(* IEC 61131-3 sources: plc-st-coding-agent/progress/evidence/f14_v14_remaining_20261113/jobs/codex_deepseek-v4pro (part 5) *)

(* ---- self-medium-04.raw_candidate_01.st ---- *)
FUNCTION_BLOCK FB
VAR_INPUT
    startBtn   : BOOL;
    resetBtn   : BOOL;
    doneSensor : BOOL;
    targetVol  : REAL;
    flowVol    : REAL;
END_VAR
VAR_OUTPUT
    valveOpen  : BOOL;
    fillsToday : INT;
END_VAR
VAR
    prevStartBtn   : BOOL := FALSE;
    prevResetBtn   : BOOL := FALSE;
    prevValveOpen  : BOOL := FALSE;
    pendingConfirm : BOOL := FALSE;
    accumulatedVol : REAL := 0.0;
    tmp_risingReset : BOOL;
    tmp_risingStart : BOOL;
    tmp_isFilling   : BOOL;
END_VAR

(* ENGINEERING_CONTRACT
   valveOpen: set only on start edge from idle/wait (R2,S2); holds while
             accumulatedVol < targetVol (R3,S9); closes on reset or target reach (R1,R3,S5).
   pendingConfirm: set same scan as target close; persists until confirmation,
             next start, or reset; sensor TRUE does not repeat count (R3-R5,S11).
   fillsToday: increments once on doneSensor with pending; saturates at 32767
             and still clears pending; reset zeros in same scan (R4-R5,S1,S6,S14).
   accumulatedVol: reset on reset/new bottle; adds flowVol only while filling,
             including start scan (R1-R3,S12).
   Priority: reset > start/new-bottle cancellation > flow/threshold close > done confirm.
   Units: targetVol/flowVol in mL REAL; fillsToday signed INT bounds 0..32767.
*)

(* CONTRACT_RULES [] *)

tmp_risingReset := resetBtn AND NOT prevResetBtn;
tmp_risingStart := startBtn AND NOT prevStartBtn;

IF tmp_risingReset THEN
    valveOpen      := FALSE;
    fillsToday     := 0;
    accumulatedVol := 0.0;
    pendingConfirm := FALSE;
ELSE
    tmp_isFilling := FALSE;

    IF tmp_risingStart AND NOT valveOpen THEN
        pendingConfirm := FALSE;
        accumulatedVol := 0.0;
        valveOpen      := TRUE;
        tmp_isFilling   := TRUE;
    ELSIF valveOpen THEN
        tmp_isFilling := TRUE;
    END_IF;

    IF tmp_isFilling THEN
        accumulatedVol := accumulatedVol + flowVol;
        IF accumulatedVol >= targetVol THEN
            valveOpen      := FALSE;
            pendingConfirm := TRUE;
            tmp_isFilling   := FALSE;
        END_IF;
    END_IF;

    IF pendingConfirm AND doneSensor THEN
        IF fillsToday < 32767 THEN
            fillsToday := fillsToday + 1;
        END_IF;
        pendingConfirm := FALSE;
    END_IF;
END_IF;

prevStartBtn  := startBtn;
prevResetBtn  := resetBtn;
prevValveOpen := valveOpen;

END_FUNCTION_BLOCK

(* ---- self-medium-05.candidate_01.st ---- *)
FUNCTION_BLOCK FB
VAR_INPUT
    enable : BOOL;
    resetBtn : BOOL;
    scanSeconds : LREAL;
    steamFlow : LREAL;
    fuelFlow : LREAL;
    steamTemp : LREAL;
    steamPressure : LREAL;
END_VAR
VAR_OUTPUT
    qualified : BOOL;
    dataFault : BOOL;
    qualifiedTon : LREAL;
    fuelTon : LREAL;
    revenue : LREAL;
    cost : LREAL;
    netProfit : LREAL;
END_VAR
VAR
    local_prev_reset : BOOL := FALSE;
    local_reset_edge : BOOL;
END_VAR

(* ENGINEERING_CONTRACT
   - qualified/dataFault: combinational, updated every scan.
   - qualifiedTon: accumulates only when enable, no fault, qualified, and no reset edge.
   - fuelTon: accumulates only when enable, no fault, and no reset edge.
   - resetBtn rising edge: clears both accumulators, higher priority than enable/fault.
   - reset is edge-only; held resetBtn does not repeatedly clear.
   - revenue/cost/netProfit recomputed every scan from current accumulators.
   - scanSeconds unit s, flows kg/s; both are legal under stated fault bounds.
*)

(* CONTRACT_RULES [] *)

local_reset_edge := resetBtn AND NOT local_prev_reset;

qualified := (steamTemp >= 447.0) AND (steamTemp <= 453.0)
             AND (steamPressure >= 3750.0) AND (steamPressure <= 3850.0);

dataFault := (scanSeconds <= 0.0)
             OR (scanSeconds > 10.0)
             OR (steamFlow < 0.0) OR (steamFlow > 90.0)
             OR (fuelFlow < 0.0) OR (fuelFlow > 6.0);

IF local_reset_edge THEN
    qualifiedTon := 0.0;
    fuelTon := 0.0;
ELSE
    IF enable AND NOT dataFault THEN
        fuelTon := fuelTon + (fuelFlow * scanSeconds / 1000.0);

        IF qualified THEN
            qualifiedTon := qualifiedTon + (steamFlow * scanSeconds / 1000.0);
        END_IF;
    END_IF;
END_IF;

revenue := qualifiedTon * 280.0;
cost := fuelTon * 1500.0;
netProfit := revenue - cost;

local_prev_reset := resetBtn;

END_FUNCTION_BLOCK

(* ---- self-medium-05.raw_candidate_01.st ---- *)
FUNCTION_BLOCK FB
VAR_INPUT
    enable : BOOL;
    resetBtn : BOOL;
    scanSeconds : LREAL;
    steamFlow : LREAL;
    fuelFlow : LREAL;
    steamTemp : LREAL;
    steamPressure : LREAL;
END_VAR
VAR_OUTPUT
    qualified : BOOL;
    dataFault : BOOL;
    qualifiedTon : LREAL;
    fuelTon : LREAL;
    revenue : LREAL;
    cost : LREAL;
    netProfit : LREAL;
END_VAR
VAR
    local_prev_reset : BOOL := FALSE;
    local_reset_edge : BOOL;
END_VAR

(* ENGINEERING_CONTRACT
   - qualified/dataFault: combinational, updated every scan.
   - qualifiedTon: accumulates only when enable, no fault, qualified, and no reset edge.
   - fuelTon: accumulates only when enable, no fault, and no reset edge.
   - resetBtn rising edge: clears both accumulators, higher priority than enable/fault.
   - reset is edge-only; held resetBtn does not repeatedly clear.
   - revenue/cost/netProfit recomputed every scan from current accumulators.
   - scanSeconds unit s, flows kg/s; both are legal under stated fault bounds.
*)

(* CONTRACT_RULES [] *)

local_reset_edge := resetBtn AND NOT local_prev_reset;

qualified := (steamTemp >= 447.0) AND (steamTemp <= 453.0)
             AND (steamPressure >= 3750.0) AND (steamPressure <= 3850.0);

dataFault := (scanSeconds <= 0.0)
             OR (scanSeconds > 10.0)
             OR (steamFlow < 0.0) OR (steamFlow > 90.0)
             OR (fuelFlow < 0.0) OR (fuelFlow > 6.0);

IF local_reset_edge THEN
    qualifiedTon := 0.0;
    fuelTon := 0.0;
ELSE
    IF enable AND NOT dataFault THEN
        fuelTon := fuelTon + (fuelFlow * scanSeconds / 1000.0);

        IF qualified THEN
            qualifiedTon := qualifiedTon + (steamFlow * scanSeconds / 1000.0);
        END_IF;
    END_IF;
END_IF;

revenue := qualifiedTon * 280.0;
cost := fuelTon * 1500.0;
netProfit := revenue - cost;

local_prev_reset := resetBtn;

END_FUNCTION_BLOCK

(* ---- self-medium-06.candidate_01.st ---- *)
FUNCTION_BLOCK FB
VAR_INPUT
    enable : BOOL;
    resetBtn : BOOL;
    sensorValid : BOOL;
    setpoint : REAL;
    temperature : REAL;
    scanSeconds : REAL;
    bias : REAL;
END_VAR
VAR_OUTPUT
    power : REAL;
    correction : REAL;
    fault : BOOL;
END_VAR
VAR
    tmp_e : REAL;
    tmp_de : REAL;
    tmp_x : REAL;
    tmp_y : REAL;
    tmp_ePrev : REAL := 0.0;
    tmp_historyValid : BOOL := FALSE;
    tmp_resetEdge : R_TRIG;
    tmp_resetPulse : BOOL;
END_VAR

(* CONTRACT_RULES [] *)

(* ENGINEERING_CONTRACT
   power: active only enable & !fault & no reset pulse; zero branch has same-scan priority; recomputed/clamped each active scan; 0..100.
   correction: computed on active scan; zero branch resets; first/cleared-history scan uses de=0; range [-30,30]; no separate clamp.
   fault: combinational from !sensorValid or scanSeconds<=0 or scanSeconds>10.
   reset: R_TRIG pulse only; held reset does not sustain zero.
   history: ePrev and historyValid retained; cleared in every zero branch; set after active computation.
   units: e degC, de degC/s, scanSeconds s, bias/power/correction %.
   derivation: 9-rule product centroid algebraically equals 20x+10y with history, 20x on first/cleared-history scan.
*)

tmp_resetEdge(CLK := resetBtn);
tmp_resetPulse := tmp_resetEdge.Q;

fault := (NOT sensorValid) OR (scanSeconds <= 0.0) OR (scanSeconds > 10.0);

IF (NOT enable) OR fault OR tmp_resetPulse THEN
    power := 0.0;
    correction := 0.0;
    tmp_ePrev := 0.0;
    tmp_historyValid := FALSE;
ELSE
    tmp_e := setpoint - temperature;

    IF NOT tmp_historyValid THEN
        tmp_de := 0.0;
    ELSE
        tmp_de := (tmp_e - tmp_ePrev) / scanSeconds;
    END_IF;

    tmp_x := LIMIT(-1.0, tmp_e / 10.0, 1.0);
    tmp_y := LIMIT(-1.0, tmp_de / 2.0, 1.0);

    IF NOT tmp_historyValid THEN
        correction := 20.0 * tmp_x;
    ELSE
        correction := 20.0 * tmp_x + 10.0 * tmp_y;
    END_IF;

    tmp_ePrev := tmp_e;
    tmp_historyValid := TRUE;

    power := LIMIT(0.0, bias + correction, 100.0);
END_IF;

END_FUNCTION_BLOCK

(* ---- self-medium-06.raw_candidate_01.st ---- *)
FUNCTION_BLOCK FB
VAR_INPUT
    enable : BOOL;
    resetBtn : BOOL;
    sensorValid : BOOL;
    setpoint : REAL;
    temperature : REAL;
    scanSeconds : REAL;
    bias : REAL;
END_VAR
VAR_OUTPUT
    power : REAL;
    correction : REAL;
    fault : BOOL;
END_VAR
VAR
    tmp_e : REAL;
    tmp_de : REAL;
    tmp_x : REAL;
    tmp_y : REAL;
    tmp_ePrev : REAL := 0.0;
    tmp_historyValid : BOOL := FALSE;
    tmp_resetEdge : R_TRIG;
    tmp_resetPulse : BOOL;
END_VAR

(* CONTRACT_RULES [] *)

(* ENGINEERING_CONTRACT
   power: active only enable & !fault & no reset pulse; zero branch has same-scan priority; recomputed/clamped each active scan; 0..100.
   correction: computed on active scan; zero branch resets; first/cleared-history scan uses de=0; range [-30,30]; no separate clamp.
   fault: combinational from !sensorValid or scanSeconds<=0 or scanSeconds>10.
   reset: R_TRIG pulse only; held reset does not sustain zero.
   history: ePrev and historyValid retained; cleared in every zero branch; set after active computation.
   units: e degC, de degC/s, scanSeconds s, bias/power/correction %.
   derivation: 9-rule product centroid algebraically equals 20x+10y with history, 20x on first/cleared-history scan.
*)

tmp_resetEdge(CLK := resetBtn);
tmp_resetPulse := tmp_resetEdge.Q;

fault := (NOT sensorValid) OR (scanSeconds <= 0.0) OR (scanSeconds > 10.0);

IF (NOT enable) OR fault OR tmp_resetPulse THEN
    power := 0.0;
    correction := 0.0;
    tmp_ePrev := 0.0;
    tmp_historyValid := FALSE;
ELSE
    tmp_e := setpoint - temperature;

    IF NOT tmp_historyValid THEN
        tmp_de := 0.0;
    ELSE
        tmp_de := (tmp_e - tmp_ePrev) / scanSeconds;
    END_IF;

    tmp_x := LIMIT(-1.0, tmp_e / 10.0, 1.0);
    tmp_y := LIMIT(-1.0, tmp_de / 2.0, 1.0);

    IF NOT tmp_historyValid THEN
        correction := 20.0 * tmp_x;
    ELSE
        correction := 20.0 * tmp_x + 10.0 * tmp_y;
    END_IF;

    tmp_ePrev := tmp_e;
    tmp_historyValid := TRUE;

    power := LIMIT(0.0, bias + correction, 100.0);
END_IF;

END_FUNCTION_BLOCK
